RoboDK station: xarm_handgesture.rdk

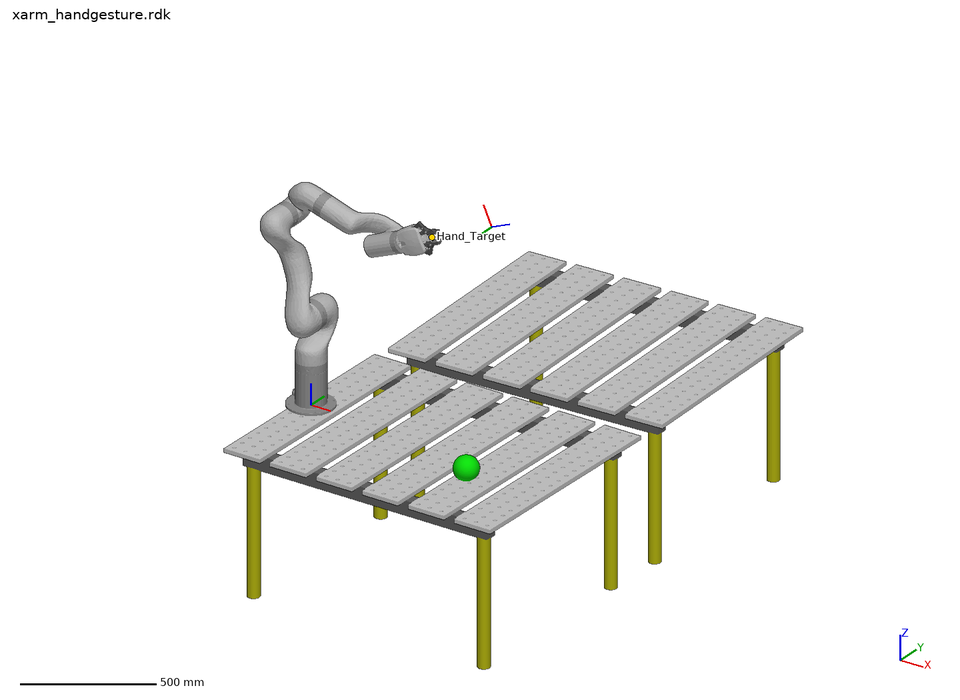
[picture v0: the station drawn from its stored meshes, robots at their saved joint values, targets as dots, program paths as lines]
Station hand_motion - Contactile (saved by RoboDK 6.0.6). Poses are relative to the parent item; angles as X-Y-Z fixed-axis rotations.
  - frame uFactory 850 Base at (0, 0, 0) mm
    - robot uFactory 850: 6 axes
        modified DH rows (alpha deg, a mm, theta deg, d mm): 0, 0, 0, 364; -90, 0, -90, 0; 0, 390, 90, 0; -90, 150, 0, 426; 90, 0, 0, 0; -90, 0, 0, 90
        joint limits [-360, -118, -225, -360, -97, -360] to [360, 120, 11, 360, 180, 360]; home [0, 0, 0, 0, 0, 0]; saved at [0.55, 18.641, -53.698, 0.823, 40.017, 1.761]
      - frame Grip_Attach_Frame at (0, -20.7, 414.56) mm
      - tool uFactory xArm Gripper, TCP at (0, 0, 140) mm, size 130.9 x 75 x 181.3 mm
    - target Hand_Target (Cartesian target) at (539.48, 3.05, 834.69) mm, rotated rx -6.31 ry -67.5 rz -173.19 deg; joints [-3.134, 2.807, -96.781, -25.954, 6.904, 29.184] of uFactory 850
    - object Sphere D100mm at (829.04, -189.85, 50.02) mm, rotated rx -179.07 ry -0.46 rz 5.2 deg, size 100 x 100 x 100 mm, geometry from Sphere-D100mm.sld
  - object Table 1200x1000mm (Welding) at (543.39, 0, 0) mm, size 1193.8 x 965.2 x 609.6 mm, geometry from Table-1200x1000mm-Welding.sld
  - object Table 1200x1000mm (Welding) at (534.06, 1058.97, 0) mm, rotated rx 0 ry 0 rz 2.59 deg, size 1193.8 x 965.2 x 609.6 mm, geometry from Table-1200x1000mm-Welding.sld
